// Generated by scripts/run_study.py. Do not edit; re-run the study instead.

FUNCTION "FC_LoadParams" : Void
TITLE = Load the designed RST and PID parameters
{ S7_Optimized_Access := 'TRUE' }
VERSION : 0.1
BEGIN
	"iRST".R[0] := 2.592645836E-01;
	"iRST".R[1] := -6.667444785E-01;
	"iRST".R[2] := 5.774055239E-01;
	"iRST".R[3] := -1.687366815E-01;
	"iRST".S[0] := 1.000000000E+00;
	"iRST".S[1] := -2.409061934E+00;
	"iRST".S[2] := 1.875383900E+00;
	"iRST".S[3] := -4.663219654E-01;
	"iRST".T[0] := 6.319795448E+01;
	"iRST".T[1] := -3.119862185E+02;
	"iRST".T[2] := 6.403125386E+02;
	"iRST".T[3] := -6.993373702E+02;
	"iRST".T[4] := 4.287036224E+02;
	"iRST".T[5] := -1.398621124E+02;
	"iRST".T[6] := 1.897277451E+01;
	"iRST".Ao[0] := 1.000000000E+00;
	"iRST".Ao[1] := -1.800000000E+00;
	"iRST".Ao[2] := 1.080000000E+00;
	"iRST".Ao[3] := -2.160000000E-01;
	"iRST".Bm[0] := 1.670439092E-03;
	"iRST".Am[0] := 1.000000000E+00;
	"iRST".Am[1] := -1.918257989E+00;
	"iRST".Am[2] := 9.199284281E-01;
	"iRST".nR := 3;
	"iRST".nS := 3;
	"iRST".nT := 6;
	"iRST".nAo := 3;
	"LineIO".PidKp := 1.083580E-01;
	"LineIO".PidTi := 4.722199E-01;
	"LineIO".PidTd := 1.686396E-01;
	"LineIO".ParamsLoaded := TRUE;
END_FUNCTION
